(* IEC 61131-3 sources: genai_codesys/experiments/raw/formal/20261109_234635_2ba96d/public_03/custom__qwen3-coder-flash/attempt_00, 2 files *)

(* ---- declaration.st ---- *)
FUNCTION_BLOCK FB_AlarmHandling
VAR_INPUT
    Value : REAL;
    hiLevel : REAL;
    loLevel : REAL;
    hystWindow : REAL;
END_VAR
VAR_OUTPUT
    hiAlarm : BOOL;
    loAlarm : BOOL;
    error : BOOL;
    status : WORD;
END_VAR

(* ---- implementation.st ---- *)
IF loLevel >= hiLevel THEN
    error := TRUE;
    status := 16#8001;
    RETURN;
END_IF;

IF hystWindow >= hiLevel - loLevel THEN
    error := TRUE;
    status := 16#8002;
    RETURN;
END_IF;

error := FALSE;
status := 16#0000;

IF Value > hiLevel THEN
    hiAlarm := TRUE;
ELSIF Value < (hiLevel - hystWindow) THEN
    hiAlarm := FALSE;
END_IF;

IF Value < loLevel THEN
    loAlarm := TRUE;
ELSIF Value > (loLevel + hystWindow) THEN
    loAlarm := FALSE;
END_IF;
